FUNCTION_BLOCK Test (* Composite Function Block Type *)
  (* Standard: 61499-2 *)
  (* Version 0.0, 7/2/2026, template *)
  PACKAGE Main;
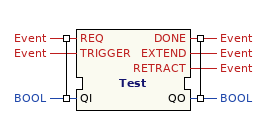
  EVENT_INPUT
    REQ WITH QI; (* Normal Execution Request *)
    TRIGGER;
  END_EVENT
  EVENT_OUTPUT
    DONE WITH QO;
    EXTEND;
    RETRACT;
  END_EVENT
  VAR_INPUT
    QI : BOOL; (* Input event qualifier *)
  END_VAR
  VAR_OUTPUT
    QO : BOOL; (* Output event qualifier *)
  END_VAR
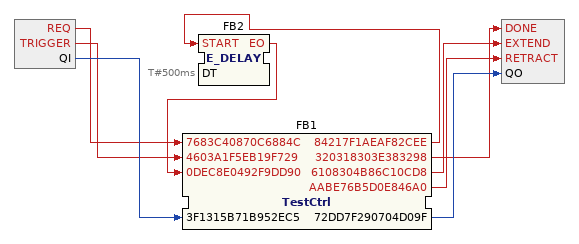
  FBS
    FB1 : TestCtrl;
    FB2 : E_DELAY(DT := T#500ms);
  END_FBS
  EVENT_CONNECTIONS
    REQ TO FB1.7683C40870C6884C;
    TRIGGER TO FB1.4603A1F5EB19F729;
    FB2.EO TO FB1.0DEC8E0492F9DD90;
    FB1.84217F1AEAF82CEE TO FB2.START;
    FB1.320318303E383298 TO DONE;
    FB1.6108304B86C10CD8 TO EXTEND;
    FB1.AABE76B5D0E846A0 TO RETRACT;
  END_CONNECTIONS
  DATA_CONNECTIONS
    QI TO FB1.3F1315B71B952EC5;
    FB1.72DD7F290704D09F TO QO;
  END_CONNECTIONS
END_FUNCTION_BLOCK
